{attribute 'qualified_only'}
VAR_GLOBAL
// 	Charger Level 1
	Inputs_1 AT%I*:ARRAY[0..19] OF BYTE;
	Outputs_1 AT%Q*:ARRAY[0..9] OF BYTE;
	
	// 	Charger Level 2
	Inputs_2 AT%I*:ARRAY[0..19] OF BYTE;
	Outputs_2 AT%Q*:ARRAY[0..9] OF BYTE;
	
	// 	Charger Level 3
	Inputs_3 AT%I*:ARRAY[0..19] OF BYTE;
	Outputs_3 AT%Q*:ARRAY[0..9] OF BYTE;
	
	// 	Charger Level 4
	Inputs_4 AT%I*:ARRAY[0..19] OF BYTE;
	Outputs_4 AT%Q*:ARRAY[0..9] OF BYTE;
	
	// 	Charger Level 5
	Inputs_5 AT%I*:ARRAY[0..19] OF BYTE;
	Outputs_5 AT%Q*:ARRAY[0..9] OF BYTE;
	
	// 	Charger Level 6
	Inputs_6 AT%I*:ARRAY[0..19] OF BYTE;
	Outputs_6 AT%Q*:ARRAY[0..9] OF BYTE;
	
	// 	Charger Level 7
	Inputs_7 AT%I*:ARRAY[0..19] OF BYTE;
	Outputs_7 AT%Q*:ARRAY[0..9] OF BYTE;
	
	// 	Charger Level 8
	Inputs_8 AT%I*:ARRAY[0..19] OF BYTE;
	Outputs_8 AT%Q*:ARRAY[0..9] OF BYTE;	
END_VAR

(* stored: Version 1.1.0.1
   GVL IO_Chargers: Id {1d018b27-eb8f-4a5e-9154-649bf0f0de30} *)
